// TIA Portal V20 export
// export: Created 2026-10-20T18:55:16.518066Z, ExportSetting None, DisplayName Totally Integrated Automation Portal, DisplayVersion V20 Update 6, DisplayName TIA Portal Openness, DisplayVersion V20 Update 6, DisplayName TIA Portal Version Control Interface, DisplayVersion V20 Update 6, DisplayName SINAMICS Startdrive Advanced, DisplayVersion V20 SP1, DisplayName SINAMICS Startdrive G130, G150, S120, S150, SINAMICS MV, G220, S200, S210, DisplayVersion V20 SP1, DisplayName SINAMICS Startdrive G110M, G120, G120C, G120D, G120P, G115D, DisplayVersion V20 SP1, DisplayName STEP 7 Professional, DisplayVersion V20 Update 6, DisplayName STEP 7 Safety, DisplayVersion V20 Update 2, DisplayName WinCC Basic/Comfort/Advanced, DisplayVersion V20 Update 6, DisplayName WinCC Unified, DisplayVersion V20 Update 6
VAR_GLOBAL   // PLC tag table "IO_Turck_4"
   "Light_Rear_1_Color1(4)" AT %QB1160 : Byte;   // Last byte - 2
   "Light_Rear_1_Intensity2(4)" AT %QB1150 : Byte;   // Last byte - 12
   "Light_Front_1_1_Direction(4)" AT %QB1112 : Byte;   // Last byte - 18
   "Light_Rear_1_Color2(4)" AT %QB1152 : Byte;   // Last byte - 10
   "Light_Rear_1_Animation(4)" AT %QB1162 : Byte;   // Last byte
   "Light_Rear_1_Percent_Width1(4)" AT %QB1146 : Byte;   // Last byte - 16
   "Light_Front_1_Percent_Width1(4)" AT %QB1114 : Byte;   // Last byte - 16
   "Light_Front_1_Speed(4)" AT %QB1124 : Byte;   // Last byte - 6
   "Light_Rear_1_Intensity1(4)" AT %QB1158 : Byte;   // Last byte - 4
   "Light_Front_1_Intensity2(4)" AT %QB1118 : Byte;   // Last byte - 12
   "Light_Rear_1_Direction(4)" AT %QB1144 : Byte;   // Last byte - 18
   "Light_Rear_1_Bounce_Style(4)" AT %QB1148 : Byte;   // Last byte - 14
   "Light_Front_1_Pulse_Pattern(4)" AT %QB1122 : Byte;   // Last byte - 8
   "Light_Front_1_Intensity1(4)" AT %QB1126 : Byte;   // Last byte - 4
   "Light_Front_1_Color2(4)" AT %QB1120 : Byte;   // Last byte - 10
   "Light_Front_1_Color1(4)" AT %QB1128 : Byte;   // Last byte - 2
   "Light_Front_1_Bounce_Style(4)" AT %QB1116 : Byte;   // Last byte - 14
   "Light_Front_1_Animation(4)" AT %QB1130 : Byte;   // Last byte
   "Light_Rear_1_Pulse_Pattern(4)" AT %QB1154 : Byte;   // Last byte - 8
   "Light_Rear_1_Speed(4)" AT %QB1156 : Byte;   // Last byte - 6
END_VAR
